(* IEC 61131-3 sources: tsplc/packages/vscode-extension/tests/fixtures/build-tool/generated/types, 7 files *)

(* ---- ST_Alarm.st ---- *)
(*
Audible alarm command for the conveyor system startup warning.
*)
TYPE ST_Alarm :
STRUCT
	(* Requests the audible startup warning. *)
	Active : BOOL;
END_STRUCT
END_TYPE

(* ---- ST_Buffer.st ---- *)
(*
Accumulation buffer capacity, occupancy count, and full status.
*)
TYPE ST_Buffer :
STRUCT
	(* Maximum occupants; zero means not configured and must inhibit admission. *)
	Capacity : UINT;
	(* FALSE until the owning PLC logic supplies a current status; FALSE on stale or unavailable inputs. *)
	Valid : BOOL;
	(* Payloads physically confirmed in this buffer. *)
	Count : UINT;
	(* Admission blocked by capacity or the configured full sensor. *)
	Full : BOOL;
END_STRUCT
END_TYPE

(* ---- ST_Button.st ---- *)
(*
Pushbutton pressed state and input validity.
*)
TYPE ST_Button :
STRUCT
	(* FALSE until the owning PLC logic supplies a current status; FALSE on stale or unavailable inputs. *)
	Valid : BOOL;
	(* TRUE while pressed; not an automatically repeating request. *)
	Pressed : BOOL;
END_STRUCT
END_TYPE

(* ---- ST_Estop.st ---- *)
(*
Supervisory emergency-stop indication for all conveyor and sorter movement. Motion requires a separate start after the stop is cleared.
*)
TYPE ST_Estop :
STRUCT
	(* FALSE until the owning PLC logic supplies a current status; FALSE on stale or unavailable inputs. *)
	Valid : BOOL;
	(* Observed global conveyor/sorter stop demand. Clearing it does not restart motion; a separate start is required. FALSE with invalid data does not indicate permission to run. *)
	Pressed : BOOL;
END_STRUCT
END_TYPE

(* ---- ST_Photoeye.st ---- *)
(*
Detection and alarm signals from a photoelectric proximity sensor.
*)
TYPE ST_Photoeye :
STRUCT
	(* Object-detection output (PNP). *)
	Detection : BOOL;
	(* Sensor alarm output. *)
	Alarm : BOOL;
END_STRUCT
END_TYPE

(* ---- ST_StackLight.st ---- *)
(*
Separate green and red lamp outputs for a two-lamp stack light. PLC logic selects the indication and times red flashing for faults.
*)
TYPE ST_StackLight :
STRUCT
	(* Switches the green lamp on when TRUE. *)
	Green : BOOL;
	(* Switches the red lamp on when TRUE; toggle in PLC logic to flash. *)
	Red : BOOL;
END_STRUCT
END_TYPE

(* ---- ST_Station.st ---- *)
(*
Operator station admission, active work, waiting queue, incoming reservations, and completed work awaiting release.
*)
TYPE ST_Station :
STRUCT
	(* Allow new admissions. Disabling does not erase existing work or reservations. *)
	Enabled : BOOL;
	(* Waiting plus incoming reservation slots; active work is separate. *)
	ReserveCapacity : UINT := 1;
	(* FALSE until the owning PLC logic supplies a current status; FALSE on stale or unavailable inputs. *)
	Valid : BOOL;
	(* Active work payload identity. *)
	ActiveId : STRING(80);
	(* Derived admission permission including QueueFull, enable, reservations, and transfer state. *)
	CanAcceptCrate : BOOL;
	(* Work completed but still physically occupies the station until outbound admission. *)
	CompletedAwaitingRelease : BOOL;
	(* Derived from configured queue sensors; do not assume suffix _1 or _2 identifies a full sensor. *)
	QueueFull : BOOL;
	(* Incoming payloads holding a waiting slot, not yet physically arrived. *)
	ReservationCount : UINT;
	(* Physically arrived waiting payloads, excluding active work and incoming reservations. *)
	WaitingCount : UINT;
END_STRUCT
END_TYPE
